SUBAPPLICATION AR_SERVER_0_1_TO_Publish_OPC (* Empfaengt einen REAL-Wert als Argument eines entfernten OPC-UA-Methodenaufrufs (CALL_METHOD, SERVER_0_1) und publiziert ihn sofort lokal weiter (PUBLISH_1) - kein VT-Anschluss, reine Weiterleitungsbruecke fuer Stationen ohne VT. Fuer 'VT-Eingabefeld auf einer anderen Station ODER Web-Dashboard rufen dieselbe Methode auf, nur bei echter Eingabe' (Franz), z.B. Druck-Referenzwerte (B20). *)
  (* Standard: 61499-2; Description: Copyright (c) 2026 Meisterschulen am Ostbahnhof This program and the accompanying materials are made available under the terms of the Eclipse Public License 2.0 which is available at https://www.eclipse.org/legal/epl-2.0/ SPDX-License-Identifier: EPL-2.0 *)
  (* Version 1.1, 2026-11-25, Franz Höpfinger, Meisterschulen am Ostbahnhof, SERVER_0_1 + E_PERMIT(PERMIT=QO) + F_MOVE(REAL) + PUBLISH_1 statt AR_SERVER_0_1/AR_PUBLISH_1: IND nur bei QO=TRUE an RSP. Ein gescheitertes RSP meldet IND mit QO=FALSE, direkt IND->RSP (in AR_SERVER_0_1) ergab eine Endlosschleife. *)
  (* Version 1.0, 2026-09-23, Franz Höpfinger, Meisterschulen am Ostbahnhof, initial implementation - Franz: 'man macht auf STG4 2 METHODEN, die werden aufgerufen: vom Web-Dashboard oder von VT1, und zwar nur wenn jemand was eingibt'. Buendelt AR_SERVER_0_1 (Empfang) + AR_PUBLISH_1 (lokale Weiterleitung), fuer Sensor-Stationen ohne eigene VT (z.B. STG4), die trotzdem echte, editierbare Referenzwerte von einer anderen Station (VT) oder dem Dashboard entgegennehmen sollen. *)
  PACKAGE MyLib::sys;
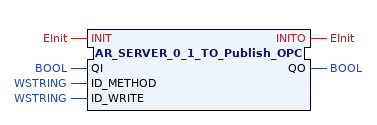
  EVENT_INPUT
    INIT : EInit; (* Initialization Request *)
  END_EVENT
  EVENT_OUTPUT
    INITO : EInit; (* Initialization Confirm *)
  END_EVENT
  VAR_INPUT
    QI : BOOL := TRUE; (* Quality Input - TRUE to enable service *)
    ID_METHOD : WSTRING; (* Lokal erzeugte OPC-UA-Methode (ACTION=CREATE_METHOD, 1 REAL-Argument) - von einer anderen Station (AR_CLIENT_1_0) UND/ODER direkt vom OPC-Dashboard aufrufbar *)
    ID_WRITE : WSTRING; (* Lokale Publish-Adresse (REAL, ACTION=PUBLISH) fuer den empfangenen Wert - typischerweise von einem lokalen Self-Subscribe gegengelesen *)
  END_VAR
  VAR_OUTPUT
    QO : BOOL; (* Quality Output - TRUE if service executed successfully *)
  END_VAR
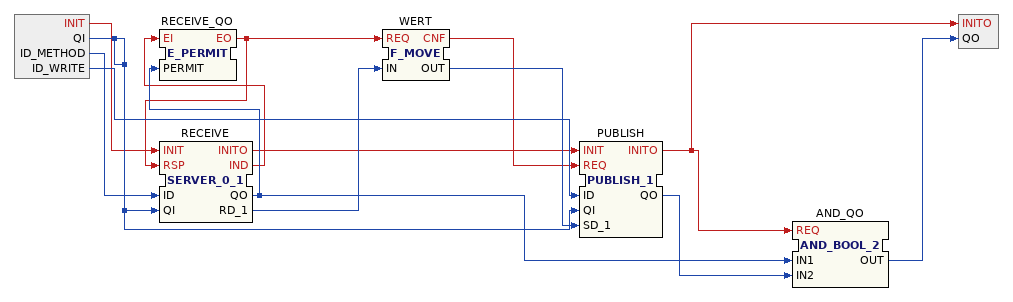
  FBS
    RECEIVE : iec61499::net::SERVER_0_1;
    RECEIVE_QO : iec61499::events::E_PERMIT; (* nur echter Call (QO=TRUE) *)
    WERT : iec61131::selection::F_MOVE; {SET_ATTRIBUTE(DataType, REAL)}
    PUBLISH : iec61499::net::PUBLISH_1;
    AND_QO : iec61131::booleanOperators::AND_BOOL_2;
  END_FBS
  EVENT_CONNECTIONS
    RECEIVE.INITO TO PUBLISH.INIT;
    INIT TO RECEIVE.INIT;
    PUBLISH.INITO TO INITO;
    PUBLISH.INITO TO AND_QO.REQ;
    RECEIVE.IND TO RECEIVE_QO.EI;
    RECEIVE_QO.EO TO RECEIVE.RSP;
    RECEIVE_QO.EO TO WERT.REQ;
    WERT.CNF TO PUBLISH.REQ;
  END_CONNECTIONS
  DATA_CONNECTIONS
    ID_METHOD TO RECEIVE.ID;
    ID_WRITE TO PUBLISH.ID;
    QI TO RECEIVE.QI;
    QI TO PUBLISH.QI;
    RECEIVE.QO TO RECEIVE_QO.PERMIT;
    RECEIVE.RD_1 TO WERT.IN;
    WERT.OUT TO PUBLISH.SD_1;
    RECEIVE.QO TO AND_QO.IN1;
    PUBLISH.QO TO AND_QO.IN2;
    AND_QO.OUT TO QO;
  END_CONNECTIONS
END_SUBAPPLICATION
